(* IEC 61131-3 sources: JingjiangMoonbox/Application/Application/任务列表/LogTask/KS_HY_日志+文件/接口功能, 5 files *)

(* ---- KS_HY_AddMsgToLog.st ---- *)
(*@CES
Name=KS_HY_AddMsgToLog
Type=FunctionBlock
TypeGuid=6f9dac99-8de1-4efc-8465-68ac443b7d08
Guid=bcb6c59b-ebd6-4321-878d-202e813fcffa
HasDeclaration=True
HasImplementation=True
*)
{DECLARATION}
FUNCTION KS_HY_AddMsgToLog : INT
(* 2025.8.23.115118
/ 添加消息到日志fifo中
*)
VAR_INPUT
	i_pstStHYLogFifo: POINTER TO StHYLogFifo;(* 日志FIFO *)
	i_iLogLevel: INT;(* 日志等级 *)
	i_sMsgContent: STRING;(* 内容部分 *)
	i_sMsgNote: STRING;(* 注解部分 *)
END_VAR
VAR
	iResult: INT;
	byIdxW_tmp: BYTE;
	pstStHYLogItem_tmp: POINTER TO StHYLogItem;
END_VAR

{IMPLEMENTATION}
iResult:= 0;
IF i_pstStHYLogFifo<>0 THEN
	(* 参数有效 *)

	(* 获取时间戳字串[YYYY/MM/DD hh:mm:ss.mmm] *)
	(* 日志内容格式:
	/ 2025/08/23 17:01:00.123[A]E-Stop Pressed.(9)
	*)
	byIdxW_tmp:= i_pstStHYLogFifo^.byIdxW;
	pstStHYLogItem_tmp:= ADR(i_pstStHYLogFifo^.astStHYLogItem[byIdxW_tmp]);
	pstStHYLogItem_tmp^.sDetails:= KS_HY_GetTimeString();

	(* 日志等级 *)
	pstStHYLogItem_tmp^.sDetails:= CONCAT(pstStHYLogItem_tmp^.sDetails, '[');
	IF i_iLogLevel=LOG_LEVEL_INFO THEN(* 一版消息 *)
		pstStHYLogItem_tmp^.sDetails:= CONCAT(pstStHYLogItem_tmp^.sDetails, 'I');
	ELSIF i_iLogLevel=LOG_LEVEL_DEBUG THEN(* 调试消息 *)
		pstStHYLogItem_tmp^.sDetails:= CONCAT(pstStHYLogItem_tmp^.sDetails, 'D');
	ELSIF i_iLogLevel=LOG_LEVEL_ALARM THEN(* 报警消息 *)
		pstStHYLogItem_tmp^.sDetails:= CONCAT(pstStHYLogItem_tmp^.sDetails, 'A');
	ELSIF i_iLogLevel=LOG_LEVEL_ERROR THEN(* 错误消息 *)
		pstStHYLogItem_tmp^.sDetails:= CONCAT(pstStHYLogItem_tmp^.sDetails, 'E');
	ELSIF i_iLogLevel=LOG_LEVEL_FATAL THEN(* 严重消息 *)
		pstStHYLogItem_tmp^.sDetails:= CONCAT(pstStHYLogItem_tmp^.sDetails, 'F');
	ELSE(* 未知消息 *)
		pstStHYLogItem_tmp^.sDetails:= CONCAT(pstStHYLogItem_tmp^.sDetails, '?');
	END_IF
	pstStHYLogItem_tmp^.sDetails:= CONCAT(pstStHYLogItem_tmp^.sDetails, ']');

	(* 日志正文 *)
	IF LEN(i_sMsgContent)>0 THEN
		pstStHYLogItem_tmp^.sDetails:= CONCAT(pstStHYLogItem_tmp^.sDetails, i_sMsgContent);
	END_IF

	(* 注解部分如果无信息/则整段不添加 *)
	IF LEN(i_sMsgNote)>0 THEN
		pstStHYLogItem_tmp^.sDetails:= CONCAT(pstStHYLogItem_tmp^.sDetails, '(');
		pstStHYLogItem_tmp^.sDetails:= CONCAT(pstStHYLogItem_tmp^.sDetails, i_sMsgNote);
		pstStHYLogItem_tmp^.sDetails:= CONCAT(pstStHYLogItem_tmp^.sDetails, ')');
	END_IF

	(* 下次写入的位置/由于接口支持多个任务调用
	/ 尽量不要直接操作i_pstStHYLogFifo内的数组索引
	*)
	byIdxW_tmp:= byIdxW_tmp+1;
	i_pstStHYLogFifo^.byIdxW:= byIdxW_tmp;
ELSE
	(* 参数无效 *)

	iResult:= -1;
END_IF

KS_HY_AddMsgToLog:= iResult;

(* ---- KS_HY_AllocGlobalMem.st ---- *)
(*@CES
Name=KS_HY_AllocGlobalMem
Type=FunctionBlock
TypeGuid=6f9dac99-8de1-4efc-8465-68ac443b7d08
Guid=11b74300-b4dc-4b42-bc03-7b37d7588a0c
HasDeclaration=True
HasImplementation=True
*)
{DECLARATION}
FUNCTION KS_HY_AllocGlobalMem : DWORD
(* 该POU建议放在系统事件PrepareStart中调用 *)
VAR_IN_OUT
	EventPrm: CmpApp.EVTPARAM_CmpApp;
END_VAR
VAR
	iResult: INT;
END_VAR

{IMPLEMENTATION}
iResult:= 0;

(* 用于文件保存时搬运的内存区域
/ 全局内存操作小于1M区域的都可以复用这个内存
*)
IF g_dwMem1MB=0 THEN
	g_dwMem1MB:= SysMemAlloc(16#100000);
END_IF

(* 火眼系统日志队列申请
/ 目前结构体中的读写索引是按照BYTE(0~255)值域覆盖范围申请数组大小的
/ 如果后续要改变数组大小/需要留意对指针索引的保护处理
*)
IF g_pstStHYLogFifo=0 THEN
	g_pstStHYLogFifo:= SysMemAlloc(SIZEOF(g_pstStHYLogFifo^));
END_IF

(* 2025.8.27.160700/han.dp
/ 增加的火眼只发数据队列内存申请
*)
IF g_pstStUdpOnlySendFifo=0 THEN
	g_pstStUdpOnlySendFifo:= SysMemAlloc(SIZEOF(g_pstStUdpOnlySendFifo^));
END_IF
KS_initStUdpOnlySendFifo(g_pstStUdpOnlySendFifo);

KS_HY_AllocGlobalMem:= INT_TO_DWORD(iResult);

(* ---- KS_HY_FileProc.st ---- *)
(*@CES
Name=KS_HY_FileProc
Type=FunctionBlock
TypeGuid=6f9dac99-8de1-4efc-8465-68ac443b7d08
Guid=f478979a-6038-403b-861a-7e2c2eb17e6a
HasDeclaration=True
HasImplementation=True
*)
{DECLARATION}
FUNCTION KS_HY_FileProc : INT
(* 火眼系统文件处理功能接口
/ ..................................................
/ 处理的文件包含两种类别: 1).系统配置参数/2).系统参数文件
/ 操作方式: AM_WRITE/AM_READ(Owner SysFile library)
/ ..................................................
/ 返回值:
/ 0.无错误/-1.传入参数非法/-2.操作的文件类型未收录
/ -3.文件访问出现错误/-4.读写的数据长度和期望的不一致
/ -5.读取的信息校验未通过/
/ -13.第2个文件写入失败
/ ..................................................
/ 特别说明:
/ 数据操作引入内存快照的原由是因为数据读写有crc校验
/ 所以在保存完成前这片内存是不能被更新的
/ 所以单独开辟了个内存区域存放一份完整的数据
*)
VAR_INPUT
	i_iFileTyp_cfg0_para1: INT;(* 0.配置信息文件/1.系统参数文件 *)
	i_xFileOpt_falseR_trueW: BOOL;(* FALSE.读操作/TRUE.写操作 *)
	i_pstStSysCfgStruct: POINTER TO StSysCfgStruct;(* 配置信息 *)
	i_pstStSysParam: POINTER TO StSysParam;(* 系统参数 *)
	i_dwDlen: DWORD;(* 数据区域大小/不包含校验 *)
	i_dwMemSnapshot: DWORD;(* 内存快照区域/系统开机就申请好1M字节/需要能涵盖保存的数据区域 *)
	i_sFileName: STRING;(* 文件名称/FNAME_SYS_CONF/FNAME_SYS_PARAM_A/FNAME_SYS_PARAM_B *)
	i_xEnableWriteFile2: BOOL;(* 使能第2个文件的写入操作/减少一次对内存的crc操作/节省时间开销 *)
	i_sFileName_2: STRING;(* 使能第2个文件的直接写入 *)
	i_pdiErrCodeEx: POINTER TO DINT;(* 返回的具体错误代码 *)
END_VAR
VAR
	iResult: INT;(* 返回值 *)

	wChk: WORD;
	dwSum: DWORD;
	wChk_tmp: WORD;
	dwSum_tmp: DWORD;

	dwDlen_AdditionInfo: DWORD;(* 附加信息长度/默认6字节/2字节CRC/4字节累加和 *)
	dwDlen_InclChk: DWORD;(* 包含校验的长度 *)
	dwDlen_Access: DWORD;(* 实际访问的有效数据长度 *)

	dwHdlFile: RTS_IEC_HANDLE;(* TYPE RTS_IEC_HANDLE : POINTER TO BYTE *)
	udiRtn: RTS_IEC_RESULT;(* TYPE RTS_IEC_RESULT : UDINT *)
						(* TYPE RTS_IEC_SIZE : POINTER TO BYTE *)
						(* RTS_INVALID_HANDLE: RTS_IEC_HANDLE(-1) *)
	rtnSFW: __XWORD;
END_VAR

{IMPLEMENTATION}
iResult:= 0;
dwDlen_AdditionInfo:= SIZEOF(wChk) + SIZEOF(dwSum);
dwDlen_InclChk:= i_dwDlen+dwDlen_AdditionInfo;
IF i_sFileName<>'' AND
	i_dwMemSnapshot<>0 AND
	(i_dwDlen>0 AND i_dwDlen<=(16#100000-dwDlen_AdditionInfo)) THEN(* 用原始参数进行判断 *)

	IF (i_iFileTyp_cfg0_para1=0 AND i_pstStSysCfgStruct<>0) OR
		(i_iFileTyp_cfg0_para1=1 AND i_pstStSysParam<>0) THEN
		(* 文件类型和其分别对应的数据地址有效 *)

		IF i_xFileOpt_falseR_trueW THEN(* 写 *)

			(* 先把内存拍照存档/之后就不用担心原数据区域发生变化了 *)
			IF i_iFileTyp_cfg0_para1=0 THEN(* 配置信息 *)
				SysMemCpy(i_dwMemSnapshot, i_pstStSysCfgStruct, i_dwDlen);
			ELSE(* 参数信息 *)
				SysMemCpy(i_dwMemSnapshot, i_pstStSysParam, i_dwDlen);
			END_IF

			(* 我们开始生成校验信息 *)
			wChk_tmp:= KS_CRC(i_dwMemSnapshot, i_dwDlen, ADR(dwSum_tmp));
			SysMemCpy(i_dwMemSnapshot+i_dwDlen, ADR(wChk_tmp), SIZEOF(wChk_tmp));
			SysMemCpy(i_dwMemSnapshot+i_dwDlen+SIZEOF(wChk_tmp), ADR(dwSum_tmp), SIZEOF(dwSum_tmp));

			(* 创建文件 *)
			dwHdlFile:= SysFileOpen(i_sFileName, SysFile.AM_WRITE, ADR(udiRtn));
			IF dwHdlFile<>RTS_INVALID_HANDLE THEN(* 成功 *)
				rtnSFW:= SysFileWrite(dwHdlFile, i_dwMemSnapshot, dwDlen_InclChk, ADR(udiRtn));
				SysFileClose(dwHdlFile);
				IF rtnSFW=0 THEN(* 写文件出现错误/曾经出现16#29(41)的错误:ERR_DISK_FULL *)

				END_IF
			ELSE(* 文件创建失败 *)
				iResult:= -3;
				IF i_pdiErrCodeEx<>0 THEN i_pdiErrCodeEx^:= UDINT_TO_DINT(udiRtn); END_IF
			END_IF

			(* 使能第2个文件写入 *)
			IF i_xEnableWriteFile2 AND
				i_sFileName_2<>'' AND
				i_sFileName_2<>i_sFileName THEN

				dwHdlFile:= SysFileOpen(i_sFileName_2, SysFile.AM_WRITE, ADR(udiRtn));
				IF dwHdlFile<>RTS_INVALID_HANDLE THEN(* 成功 *)
					rtnSFW:= SysFileWrite(dwHdlFile, i_dwMemSnapshot, dwDlen_InclChk, ADR(udiRtn));
					SysFileClose(dwHdlFile);
					IF rtnSFW=0 THEN(* 写文件出现错误/曾经出现16#29(41)的错误:ERR_DISK_FULL *)

					END_IF
				ELSE(* 文件创建失败 *)
					iResult:= -13;
					IF i_pdiErrCodeEx<>0 THEN i_pdiErrCodeEx^:= UDINT_TO_DINT(udiRtn); END_IF
				END_IF
			END_IF

		ELSE(* 读 *)

			(* 打开文件 *)
			dwHdlFile:= SysFileOpen(i_sFileName, SysFile.AM_READ, ADR(udiRtn));
			IF dwHdlFile<>RTS_INVALID_HANDLE THEN(* 成功 *)

				(* 搬运到内存后就尽快关闭文件 *)
				dwDlen_Access:= SysFileRead(dwHdlFile, i_dwMemSnapshot, dwDlen_InclChk, ADR(udiRtn));
				SysFileClose(dwHdlFile);

				(* 开始进行内存的操作 *)
				IF dwDlen_Access=dwDlen_InclChk THEN(* 数据量有效 *)

					(* 先把文件保存的校验信息读取出来 *)
					SysMemCpy(ADR(wChk), i_dwMemSnapshot+i_dwDlen, SIZEOF(wChk));
					SysMemCpy(ADR(dwSum), i_dwMemSnapshot+i_dwDlen+SIZEOF(wChk), SIZEOF(dwSum));

					(* 我们再复算一遍校验信息 *)
					wChk_tmp:= KS_CRC(i_dwMemSnapshot, i_dwDlen, ADR(dwSum_tmp));

//2026.4.6.122232增加累加和不为0
					IF wChk=wChk_tmp AND dwSum=dwSum_tmp AND dwSum<>0 THEN(* 校验信息通过 *)

						(* 可以直接搬运到目标内存区域 *)
						IF i_iFileTyp_cfg0_para1=0 THEN
							SysMemCpy(i_pstStSysCfgStruct, i_dwMemSnapshot, i_dwDlen);
						ELSE
							SysMemCpy(i_pstStSysParam, i_dwMemSnapshot, i_dwDlen);
						END_IF
					ELSE
						iResult:= -5;
					END_IF
				ELSE(* 数据量不足或者读取时出现错误 *)
					iResult:= -4;
					IF i_pdiErrCodeEx<>0 THEN i_pdiErrCodeEx^:= UDINT_TO_DINT(udiRtn); END_IF
				END_IF
			ELSE(* 文件打开失败 *)
				iResult:= -3;
				IF i_pdiErrCodeEx<>0 THEN i_pdiErrCodeEx^:= UDINT_TO_DINT(udiRtn); END_IF
			END_IF
		END_IF
	ELSE
		iResult:= -2;
	END_IF
ELSE
	iResult:= -1;
END_IF

KS_HY_FileProc:= iResult;

(* ---- KS_HY_GetTimeString.st ---- *)
(*@CES
Name=KS_HY_GetTimeString
Type=FunctionBlock
TypeGuid=6f9dac99-8de1-4efc-8465-68ac443b7d08
Guid=6552801a-dd25-4c90-9866-0e8db1fb41da
HasDeclaration=True
HasImplementation=True
*)
{DECLARATION}
FUNCTION KS_HY_GetTimeString : STRING
VAR_INPUT
END_VAR
VAR
	sFinal: STRING;
	udiResult: RTS_IEC_RESULT;
	stUTC_Timestamp: SysTime;
	stdNow: SysTimeDate;
	s_year: STRING;
	s_month: STRING;
	s_day: STRING;
	s_hour: STRING;
	s_minute: STRING;
	s_second: STRING;
	s_milliseconds: STRING;
(* 保留效率测试的部分痕迹
	stUTC_Timestamp_2: SysTime;
	ulElapsed: ULINT;
*)
END_VAR

{IMPLEMENTATION}
(* 获取时间戳字串 *)
udiResult:= SysTimeRtcHighResGet(stUTC_Timestamp);
udiResult:= SysTimeRtcConvertHighResToLocal(stUTC_Timestamp, stdNow);

s_year:=
KS_HY_UINT_TO_STRING(stdNow.wYear, 4);

s_month:=
KS_HY_UINT_TO_STRING(stdNow.wMonth, 2);

s_day:=
KS_HY_UINT_TO_STRING(stdNow.wDay, 2);

s_hour:=
KS_HY_UINT_TO_STRING(stdNow.wHour, 2);

s_minute:=
KS_HY_UINT_TO_STRING(stdNow.wMinute, 2);

s_second:=
KS_HY_UINT_TO_STRING(stdNow.wSecond, 2);

s_milliseconds:=
KS_HY_UINT_TO_STRING(stdNow.wMilliseconds, 3);

sFinal:= s_year;
sFinal:= CONCAT(sFinal, '/');
sFinal:= CONCAT(sFinal, s_month);
sFinal:= CONCAT(sFinal, '/');
sFinal:= CONCAT(sFinal, s_day);
sFinal:= CONCAT(sFinal, ' ');
sFinal:= CONCAT(sFinal, s_hour);
sFinal:= CONCAT(sFinal, ':');
sFinal:= CONCAT(sFinal, s_minute);
sFinal:= CONCAT(sFinal, ':');
sFinal:= CONCAT(sFinal, s_second);
sFinal:= CONCAT(sFinal, '.');
sFinal:= CONCAT(sFinal, s_milliseconds);

(*实测字符串操作耗时远远小于1ms
Result:= SysTimeRtcHighResGet(stUTC_Timestamp_2);
ulElapsed:= stUTC_Timestamp_2-stUTC_Timestamp;
*)

KS_HY_GetTimeString:= sFinal;

(* ---- KS_HY_UINT_TO_STRING.st ---- *)
(*@CES
Name=KS_HY_UINT_TO_STRING
Type=FunctionBlock
TypeGuid=6f9dac99-8de1-4efc-8465-68ac443b7d08
Guid=e624a904-2250-46e3-9cf7-e5a73eed6aa1
HasDeclaration=True
HasImplementation=True
*)
{DECLARATION}
FUNCTION KS_HY_UINT_TO_STRING : STRING
VAR_INPUT
	i_uiNum: UINT;(* 传入数值 *)
	i_uiLen_fixedwidth: UINT;(* 固定长度 *)
END_VAR
VAR
	uiN: UINT;
	sPrefix: STRING := '0';
	sResult: STRING := '';
	sTmp_raw: STRING := '';
	uiLen_raw: UINT;
END_VAR

{IMPLEMENTATION}
IF i_uiLen_fixedwidth>0 THEN
	sTmp_raw:= UINT_TO_STRING(i_uiNum);(* 原始数值直接转STRING *)
	uiLen_raw:= UDINT_TO_UINT(LEN(sTmp_raw));(* 看转换后长度是否满足 *)
	IF uiLen_raw>i_uiLen_fixedwidth THEN(* 原始数据超过了宽度 *)
		sResult:= MID(sTmp_raw, i_uiLen_fixedwidth, uiLen_raw-i_uiLen_fixedwidth+1);
	ELSIF uiLen_raw<i_uiLen_fixedwidth THEN(* 原始数据不够宽度 *)
		FOR uiN:=1 TO (i_uiLen_fixedwidth-uiLen_raw) BY 1 DO
			sResult:= CONCAT(sResult, sPrefix);
		END_FOR
		sResult:= CONCAT(sResult, sTmp_raw);
	ELSE(* 宽度匹配 *)
		sResult:= sTmp_raw;
	END_IF
END_IF

KS_HY_UINT_TO_STRING:= sResult;
